(* CODESYS project plcresponse.library
   DefaultNamespace: KOSTAL.TC3.Core.plcResponse
   Description: Data type for responses of PLC procedures that will result in pass or fail.
   Author: Frank Dümpelmann
   DocFormat: reStructuredText
   Title: KOSTAL.TC3.Core.plcResponse
   Version: 2019.1.0.0
   Company: KOSTAL GmbH & Co.KG
   Placeholder: KOSTAL.TC3.Core.plcResponse

Project tree, tasks and I/O mapping:
  libraries: KOSTAL.TC3.Core.functionResponse, 2019.1.0.0 (KOSTAL GmbH & Co.KG); KOSTAL.TC3.Core.process, 2019.5.0.0 (KOSTAL GmbH & Co.KG); KOSTAL.TC3.Core.Settings, 2019.0.1.0 (KOSTAL GmbH & Co.KG); KOSTAL.TC3.Components.ListOf.Objects, 2019.1.0.0 (KOSTAL GmbH & Co.KG); KOSTAL.TC3.Core.System, 2019.0.0.0 (KOSTAL GmbH & Co.KG)
  DUT/
    ListOf/
      function block FB_ListOf_PlcResponse [ST]: _deletePayLoad, _Get_P, _New, Add_DUT, CopyFrom, CopyTo, Delete_DUT, Get_I, Get_IOwner
      interface I_ListOf_PlcResponse: CopyTo, Get_I
      interface I_ListOf_PlcResponse_CopyFrom: CopyFrom
      interface I_ListOf_PlcResponse_Owner: Add_DUT, CopyFrom, CopyTo, Delete_DUT, Get_I, Get_IOwner
    function block FB_PlcResponse [ST]: clear, CopyFrom, description, fail, pass
    interface I_plcResponse: description, fail, pass
    interface I_plcResponse_Owner: description, fail, pass
  Project Information/
    function F_GetCompany [ST]
    function F_GetTitle [ST]
    function F_GetVersion [ST]
  Version/
    global variables Global_Version
*)

// Version/Global_Version
{attribute 'TcGenerated'}
{attribute 'no-analysis'}
{attribute 'linkalways'}
// This function has been automatically generated from the project information.
VAR_GLOBAL CONSTANT
	{attribute 'const_non_replaced'}
	stLibVersion_KOSTAL_TC3_Core_plcResponse : ST_LibVersion := (iMajor := 2019, iMinor := 1, iBuild := 0, iRevision := 0, nFlags := 1, sVersion := '2019.1.0.0');
END_VAR

// DUT/ListOf/FB_ListOf_PlcResponse
FUNCTION_BLOCK FB_ListOf_PlcResponse  EXTENDS KOSTAL_TC3_Components_ListOf_Objects.FB_Base IMPLEMENTS I_ListOf_PlcResponse, I_ListOf_PlcResponse_CopyFrom, I_ListOf_PlcResponse_Owner

VAR
	_Dummy	: FB_PlcResponse;
END_VAR

//Overwrites the method in the base class with the real contents of the ListOf class.
METHOD PROTECTED  _deletePayLoad
VAR_INPUT
	pPayload	:	PVOID; 
END_VAR

VAR
	_p	: POINTER TO FB_PlcResponse;
END_VAR

IF pPayload = 0  THEN	RETURN;	END_IF

_p:= pPayload;

__DELETE(_p);
END_METHOD

//Get read/write access to content
//Get_P returns a pointer to the Dummy instance
METHOD PROTECTED _Get_P : POINTER TO FB_PlcResponse

VAR_INPUT
	NumberOfObject	: UDINT;
	Response				: REFERENCE TO KOSTAL_TC3_Core_functionResponse.FB_functionResponse;
END_VAR

VAR
	_response: KOSTAL_TC3_Core_functionResponse.FB_functionResponse;
END_VAR

_response.clear();

IF (NumberOfObject = 0) 
OR (NumberOfObject > _ListOfObject.nObjects)
OR (_ListOfObject.pObjects = 0)
THEN

	_Dummy.Clear();

	_Get_P:= ADR(_Dummy);

	_response.status:= 'return Dummy because NumberOfPosition is out of range';

ELSE

	_response.success:= TRUE;
	
	_Get_P:= _ListOfObject.pObjects[NumberOfObject - 1];

END_IF

IF __ISVALIDREF(Response) THEN	Response.CopyFrom(_response);	END_IF
END_METHOD

//Overwrites the method in the base class with the real contents of the ListOf class.
METHOD PROTECTED  _New : PVOID

VAR
	_pNew: POINTER TO FB_PlcResponse;
END_VAR

_pNew:= __NEW(FB_PlcResponse);

_New:= _pNew;
END_METHOD

//Add a new instance of FB_Dut and copy content from [IN] to the new instance
METHOD PUBLIC Add_DUT : BOOL
VAR_INPUT
	IN				: I_PlcResponse;
	Response	: REFERENCE TO KOSTAL_TC3_Core_functionResponse.FB_functionResponse;
END_VAR

VAR
	pDUT: POINTER TO FB_PlcResponse;
	_response: KOSTAL_TC3_Core_functionResponse.FB_functionResponse;
END_VAR
_response.clear();

//create a new empty object 
IF NOT _AddObject() THEN
	_response.status:= ('_AddObject failed');
	IF __ISVALIDREF(Response) THEN	Response.CopyFrom(_response);	END_IF
	RETURN;	
END_IF

//Return, if no  [IN] object is available
IF IN = 0 THEN 
	_response.status:= ('IN Parameter not defined');
	IF __ISVALIDREF(Response) THEN	Response.CopyFrom(_response);	END_IF
	RETURN;	
END_IF

//otherwise fill [IN] object content to new virtual instance
pDUT:= _Get_P(_ListOfObject.nObjects, _response);

IF NOT _response.success THEN 
	IF __ISVALIDREF(Response) THEN	Response.CopyFrom(_response);	END_IF
	RETURN;	
END_IF

IF pDUT = 0 THEN 
	_response.status:= ('no Pointer get from list');
	IF __ISVALIDREF(Response) THEN	Response.CopyFrom(_response);	END_IF
	RETURN;	
END_IF

pDut^.CopyFrom(IN);

_response.success:= TRUE;
IF __ISVALIDREF(Response) THEN	Response.CopyFrom(_response);	END_IF

Add_DUT:= TRUE;
END_METHOD

METHOD PUBLIC CopyFrom
VAR_INPUT
	IN	: I_ListOf_PlcResponse;
END_VAR

VAR
	_udi: UDINT;
END_VAR

IF IN = 0 THEN RETURN;	END_IF

Clear();

FOR _udi:= 1 TO IN.NumberOfObjects DO
	Add_DUT(IN.Get_I(_udi, 0), 0);
END_FOR
END_METHOD

METHOD PUBLIC CopyTo
VAR_INPUT
	IN	: I_ListOf_PlcResponse_CopyFrom;
END_VAR

IF IN = 0 THEN RETURN;	END_IF

IN.CopyFrom(THIS^);
END_METHOD

METHOD PUBLIC Delete_DUT : BOOL
VAR_INPUT
	Number	: UDINT;	//Number of DUT in List
END_VAR

VAR
	_Set: FB_ListOf_PlcResponse;
	_udi: UDINT;
END_VAR

//Range control
IF Number = 0 							THEN RETURN;	END_IF
IF Number > NumberOfObjects	THEN RETURN;	END_IF

//Intermediate storage - prepare
_Set.Clear();

//catch all elements without the Number defiend
FOR _udi:= 1 TO NumberOfObjects DO
	IF _udi <> Number THEN
		_Set.Add_DUT(THIS^.Get_I(_udi, 0), 0);
	END_IF
END_FOR

//Delete own content
Clear();

//Add the remaining elements of the own class. 
FOR _udi:= 1 TO _Set.NumberOfObjects DO
		THIS^.Add_DUT(_Set.Get_I(_udi, 0), 0);
END_FOR

//Intermediate storage - clean Router storage
_Set.Clear();

Delete_DUT:= TRUE;
END_METHOD

//Get readonly access to content 
METHOD Get_I : I_PlcResponse

VAR_INPUT
	NumberOfObject	: UDINT;
	Response				: REFERENCE TO KOSTAL_TC3_Core_functionResponse.FB_functionResponse;
END_VAR

VAR
	_response: KOSTAL_TC3_Core_functionResponse.FB_functionResponse;
END_VAR

_response.clear();

Get_I:= _Get_P(NumberOfObject, _response)^;

IF __ISVALIDREF(Response) THEN	Response.CopyFrom(_response);	END_IF
END_METHOD

//Get full access to content 
METHOD Get_IOwner : I_PlcResponse_Owner

VAR_INPUT
	NumberOfObject	: UDINT;
	Response				: REFERENCE TO KOSTAL_TC3_Core_functionResponse.FB_functionResponse;
END_VAR

VAR
	_response: KOSTAL_TC3_Core_functionResponse.FB_functionResponse;
END_VAR

_response.clear();

Get_IOwner:= _Get_P(NumberOfObject, _response)^;

IF __ISVALIDREF(Response) THEN	Response.CopyFrom(_response);	END_IF
END_METHOD

END_FUNCTION_BLOCK

// DUT/ListOf/I_ListOf_PlcResponse
INTERFACE I_ListOf_PlcResponse EXTENDS KOSTAL_TC3_Components_ListOf_Objects.I_Base

METHOD PUBLIC CopyTo
VAR_INPUT
	IN	: I_ListOf_PlcResponse_CopyFrom;
END_VAR
END_METHOD

METHOD Get_I : I_PlcResponse

VAR_INPUT
	NumberOfObject	: UDINT;
	Response				: REFERENCE TO KOSTAL_TC3_Core_functionResponse.FB_functionResponse;
END_VAR
END_METHOD

END_INTERFACE

// DUT/ListOf/I_ListOf_PlcResponse_CopyFrom
INTERFACE I_ListOf_PlcResponse_CopyFrom EXTENDS KOSTAL_TC3_Core_System.I_Interface

METHOD PUBLIC CopyFrom
VAR_INPUT
	IN	: I_ListOf_PlcResponse;
END_VAR
END_METHOD

END_INTERFACE

// DUT/I_plcResponse
INTERFACE I_plcResponse EXTENDS KOSTAL_TC3_Core_process.I_processState

PROPERTY PUBLIC description : KOSTAL_TC3_Core_Settings.T_MaxString
GET
END_GET
END_PROPERTY

PROPERTY PUBLIC fail : BOOL
GET
END_GET
END_PROPERTY

PROPERTY PUBLIC pass : BOOL
GET
END_GET
END_PROPERTY

END_INTERFACE

// DUT/ListOf/I_ListOf_PlcResponse_Owner
INTERFACE I_ListOf_PlcResponse_Owner EXTENDS KOSTAL_TC3_Components_ListOf_Objects.I_Base_Owner

//Add a new instance of FB_Dut and copy content from [IN] to the new instance
METHOD PUBLIC Add_DUT : BOOL
VAR_INPUT
	IN				: I_PlcResponse;
	Response	: REFERENCE TO KOSTAL_TC3_Core_functionResponse.FB_functionResponse;
END_VAR
END_METHOD

METHOD PUBLIC CopyFrom
VAR_INPUT
	IN	: I_ListOf_PlcResponse;
END_VAR
END_METHOD

METHOD PUBLIC CopyTo
VAR_INPUT
	IN	: I_ListOf_PlcResponse_CopyFrom;
END_VAR
END_METHOD

METHOD PUBLIC Delete_DUT : BOOL
VAR_INPUT
	Number	: UDINT;	//Number of DUT in List
END_VAR
END_METHOD

//Get readonly access to content 
METHOD Get_I : I_PlcResponse

VAR_INPUT
	NumberOfObject	: UDINT;
	Response				: REFERENCE TO KOSTAL_TC3_Core_functionResponse.FB_functionResponse;
END_VAR
END_METHOD

//Get full access to content 
METHOD Get_IOwner : I_PlcResponse_Owner

VAR_INPUT
	NumberOfObject	: UDINT;
	Response				: REFERENCE TO KOSTAL_TC3_Core_functionResponse.FB_functionResponse;
END_VAR
END_METHOD

END_INTERFACE

// DUT/I_plcResponse_Owner
INTERFACE I_plcResponse_Owner EXTENDS KOSTAL_TC3_Core_process.I_processState_Owner

PROPERTY PUBLIC description : KOSTAL_TC3_Core_Settings.T_MaxString
GET
END_GET
SET
END_SET
END_PROPERTY

PROPERTY PUBLIC fail : BOOL
GET
END_GET
SET
END_SET
END_PROPERTY

PROPERTY PUBLIC pass : BOOL
GET
END_GET
SET
END_SET
END_PROPERTY

END_INTERFACE

// DUT/FB_PlcResponse
(*

:Author: Frank Dümpelmann <f.duempelmann@kostal.com>
:Date: 2018-10-26

Function
========
Data type for responses of PLC procedures that will result in pass or fail.

Methods and Properties
======================
| pass 		:BOOL 	PLC procedure sucessfully finished
| fail		:BOOL 	PLC procedure failde
| status	:STRING Fault description in case of failure
| clear()	METHOD	Reset all values

*)

{attribute 'enable_dynamic_creation'}
FUNCTION_BLOCK PUBLIC FB_PlcResponse EXTENDS KOSTAL_TC3_Core_process.FB_processState IMPLEMENTS I_plcResponse, I_plcResponse_Owner

VAR
	_pass					: BOOL;
	_fail					: BOOL;
	_description	: KOSTAL_TC3_Core_Settings.T_MaxString;
END_VAR

METHOD PUBLIC clear

SUPER^.clear();

_pass:= FALSE;
_fail:= FALSE;

_description:= '';
END_METHOD

METHOD PUBLIC CopyFrom
VAR_INPUT
	IN	: I_processState;
END_VAR

VAR
	_obj	: I_plcResponse;
	_bResult: BOOL;
END_VAR

IF IN = 0 THEN	RETURN;	END_IF

_bResult := __QUERYINTERFACE(IN, _obj);
 
IF NOT _bResult THEN RETURN;	END_IF
IF _obj = 0 THEN RETURN;	END_IF

SUPER^.CopyFrom(IN);
_pass					:= _obj.pass;
_fail					:= _obj.fail;
_description	:= _obj.description;
END_METHOD

PROPERTY PUBLIC description : KOSTAL_TC3_Core_Settings.T_MaxString
GET

description:= _description;
END_GET
SET

_description:= description;
END_SET
END_PROPERTY

PROPERTY PUBLIC fail : BOOL
GET

fail:= _fail;
END_GET
SET

_fail:= fail;
END_SET
END_PROPERTY

PROPERTY PUBLIC pass : BOOL
GET

pass:= _pass;
END_GET
SET

_pass:= pass;
END_SET
END_PROPERTY

END_FUNCTION_BLOCK

// Project Information/F_GetCompany
// This function has been automatically generated from the project information.
{attribute 'signature_flag' := '1073741824'}
{attribute 'TcGenerated'}
{attribute 'no-analysis'}
FUNCTION F_GetCompany : WSTRING
VAR_INPUT
	
END_VAR

F_GetCompany := "KOSTAL GmbH & Co.KG";

END_FUNCTION

// Project Information/F_GetTitle
// This function has been automatically generated from the project information.
{attribute 'signature_flag' := '1073741824'}
{attribute 'TcGenerated'}
{attribute 'no-analysis'}
FUNCTION F_GetTitle : WSTRING
VAR_INPUT
	
END_VAR

F_GetTitle := "KOSTAL.TC3.Core.plcResponse";

END_FUNCTION

// Project Information/F_GetVersion
// This function has been automatically generated from the project information.
{attribute 'signature_flag' := '1073741824'}
{attribute 'TcGenerated'}
{attribute 'no-analysis'}
FUNCTION F_GetVersion : ST_LibVersion
VAR_INPUT
	
END_VAR

F_GetVersion.iMajor := 2019;
F_GetVersion.iMinor := 1;
F_GetVersion.iBuild := 0;
F_GetVersion.iRevision := 0;
F_GetVersion.sVersion := '2019.1.0.0';
F_GetVersion.nFlags := 1;

END_FUNCTION
